(* IEC 61131-3 sources: Caravan/Archiv/12-04-19/Stations/MachineControl/MachineControl/Class/NightLight_Class, 1 file *)

(* ---- NightLight_Class.st ---- *)
(*!
<Class
	Name               = "NightLight_Class"
	Revision           = "0.0"
	RealtimeTask       = "false"
	CyclicTask         = "true"
	DefCyclictime      = "50 µs"
	BackgroundTask     = "false"
	Sigmatek           = "false"
	OSInterface        = "false"
	HighPriority       = "false"
	Automatic          = "false"
	UpdateMode         = "Prescan"
	SharedCommandTable = "true"
	Objectsize         = "(780,180)">
	<Channels>
		<Server Name="ClassSvr" Visualized="false" Initialize="false" WriteProtected="true" Retentive="false"/>
		<Server Name="NightlightHZS_S" Visualized="true" Remotely="true" Initialize="false" WriteProtected="false" Retentive="false"/>
		<Server Name="sBrightness" Visualized="true" Initialize="true" DefValue="0" WriteProtected="false" Retentive="SRam"/>
		<Client Name="cNightlightSwitch" Required="true" Internal="false"/>
		<Client Name="OC_To_Timer_Class" Required="true" Internal="false"/>
	</Channels>
</Class>
*)
NightLight_Class : CLASS
  //Servers:
	ClassSvr 	: SvrChCmd_DINT;
	NightlightHZS_S 	: SvrCh_DINT;
	sBrightness 	: SvrCh_DINT;
  //Clients:
	OC_To_Timer_Class 	: CltChCmd_Timer_Class;
	cNightlightSwitch 	: CltCh_DINT;
  //Variables:
  //Functions:

	FUNCTION VIRTUAL GLOBAL CyWork
		VAR_INPUT
			EAX 	: UDINT;
		END_VAR
		VAR_OUTPUT
			state (EAX) 	: UDINT;
		END_VAR;
  //Tables:
	FUNCTION @STD
		VAR_OUTPUT
			ret_code	: CONFSTATES;
		END_VAR;
	FUNCTION GLOBAL TAB @CT_;
END_CLASS;

#pragma usingLtd Timer_Class

FUNCTION VIRTUAL GLOBAL NightLight_Class::CyWork
	VAR_INPUT
		EAX 	: UDINT;
	END_VAR
	VAR_OUTPUT
		state (EAX) 	: UDINT;
	END_VAR

  //Read

  cNightlightSwitch :=  cNightlightSwitch.Read();

  NightlightHZS_S   :=   NightlightHZS_S.Read();

  sBrightness       :=   sBrightness.Read();

  if OC_To_Timer_Class.Nachtmodus_S = 1 & NightlightHZS_S = 1 then

        cNightlightSwitch   :=    cNightlightSwitch.Write(input:=sBrightness);

     else

        cNightlightSwitch   :=    cNightlightSwitch.Write(input:=0);

  end_if;

	state := READY;

END_FUNCTION
